// TIA Portal V21 export
// export: Created 2026-11-21T13:54:31.1489017Z, ExportSetting WithDefaults, DisplayName Totally Integrated Automation Portal, DisplayVersion V21, DisplayName STEP 7 Professional, DisplayVersion V21, DisplayName STEP 7 Safety, DisplayVersion V21, DisplayName Tech WebApplication, DisplayVersion V21, DisplayName WinCC Basic/Comfort/Advanced, DisplayVersion V21, DisplayName WinCC Unified, DisplayVersion V21
Screen "Pump"  1024x768, Number=2
  ScreenLayer 
    TextField "SpeedLabel" at 20,40 size 160x30  StyleItem=Text field, Text="Pump speed"
    IOField "SpeedValue" at 200,40 size 120x30  DataFormat=Decimal, FormatPattern=999.999, Mode=InOutput, StyleItem=I/O field
